(* PLC project v0.5.3_PreCommissioningPrep.project, CODESYS CODESYS V3.5 SP19 Patch 1 *)
(* stored: creationDateTime 2026-07-30T00:34:09.1408011, modificationDateTime 2026-07-28T11:53:41.5518987 *)

PROGRAM POU
  VAR
    instInput00 : FB_INPUT;
    instJoystick01 : FB_JOYSTICK;
    instSafetyM1 : FB_SAFETY_WINCH;
  END_VAR

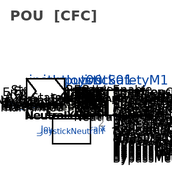
(* CFC diagram, written out as Structured Text *)
instInput00(InputRaw := M1_BrakeIsOpen_DI);
instJoystick01(Enable := instInput00.State, NeutralXMem := _JoystickNeutralX, NeutralYMem := _JoystickNeutralY);
instSafetyM1(Enable := instJoystick01.Ready);
END_PROGRAM
